Fanuc KAREL source: kt00206.KL

-- PROVISIONAL review KL for V770-1; original PC SHA256 3de2cc6922501834d98956aaef8b2fe474f1a10a44e0f9b797e71d65658a5f7a
-- Incomplete behavior may be omitted. Consult companion uncertainty JSON. Do not deploy.
PROGRAM KT00206
%NOLOCKGROUP
VAR
  I1 : INTEGER
  OUT : INTEGER
-- UNRESOLVED_DECL Y2 type=002018
BEGIN
  -- UNRESOLVED_PC offsets 5-16; opcodes 2E,23
  -- UNRESOLVED_PC offsets 21-35; opcodes 2E,22,9D,33,B2
  -- UNRESOLVED_PC offsets 40-62; opcodes 21,22,9D,33,B1,46,23
  -- UNRESOLVED_PC offsets 67-71; opcodes 7F
END KT00206
